// Minimal I_Comm stub for tests: every Publish/PublishLog call is a no-op that reports success,
// so FBs under test can call fbComm.Publish(...) freely without a real MQTT connection.
FUNCTION_BLOCK FB_NullComm IMPLEMENTS BROTLib.I_Comm
VAR
END_VAR

METHOD Publish : BOOL
VAR_INPUT
	domain			: STRING(255) := 'environment';
	location		: STRING(255) := 'roof';
	parameter		: STRING(255);
	value			: STRING(255);
END_VAR
VAR_OUTPUT
	published	: BOOL;
END_VAR
Publish := TRUE;
published := TRUE;
END_METHOD

METHOD PublishLREAL : BOOL
VAR_INPUT
	domain			: STRING(255) := 'environment';
	location		: STRING(255) := 'roof';
	parameter		: STRING(255);
	value			: LREAL;
END_VAR
VAR_OUTPUT
	published	: BOOL;
END_VAR
PublishLREAL := TRUE;
published := TRUE;
END_METHOD

METHOD PublishINT : BOOL
VAR_INPUT
	domain			: STRING(255) := 'environment';
	location		: STRING(255) := 'roof';
	parameter		: STRING(255);
	value			: LINT;
END_VAR
VAR_OUTPUT
	published	: BOOL;
END_VAR
PublishINT := TRUE;
published := TRUE;
END_METHOD

METHOD PublishBOOL : BOOL
VAR_INPUT
	domain			: STRING(255) := 'environment';
	location		: STRING(255) := 'roof';
	parameter		: STRING(255);
	value			: BOOL;
END_VAR
VAR_OUTPUT
	published	: BOOL;
END_VAR
PublishBOOL := TRUE;
published := TRUE;
END_METHOD

METHOD PublishString : BOOL
VAR_INPUT
	domain			: STRING(255) := 'environment';
	location		: STRING(255) := 'roof';
	parameter		: STRING(255);
	value			: STRING(255);
END_VAR
VAR_OUTPUT
	published	: BOOL;
END_VAR
PublishString := TRUE;
published := TRUE;
END_METHOD

METHOD PublishLog : BOOL
VAR_INPUT
	level		: STRING(255) := 'INFO';
	message		: STRING(255);
END_VAR
VAR_OUTPUT
	published	: BOOL;
END_VAR
PublishLog := TRUE;
published := TRUE;
END_METHOD

END_FUNCTION_BLOCK

(* stored: Version 1.1.0.1, ProductVersion 3.1.4024.15
   POU FB_NullComm: Id {74fa3d1a-677d-5009-aa28-dee94c7877db}, SpecialFunc None
   Method Publish: Id {f28635a0-98ee-5d5d-8fa2-ab05dd592243}
   Method PublishLREAL: Id {32399ef0-2ca1-57e7-95eb-1a6bb9ed7608}
   Method PublishINT: Id {5985129e-f1f9-5c2c-960b-660bc2fac4ec}
   Method PublishBOOL: Id {3b55248f-9707-5979-880f-812b2bad7d79}
   Method PublishString: Id {bbe9bc8d-29ad-58c3-8713-b5201422cb32}
   Method PublishLog: Id {bba6b9a2-4491-5f6d-b181-ac9167d5e786} *)
